// TIA Portal V21 export
// export: Created 2026-11-07T17:04:58.8890969Z, ExportSetting WithDefaults, DisplayName Totally Integrated Automation Portal, DisplayVersion V21, DisplayName STEP 7 Professional, DisplayVersion V21, DisplayName STEP 7 Safety, DisplayVersion V21, DisplayName Tech WebApplication, DisplayVersion V21, DisplayName WinCC Basic/Comfort/Advanced, DisplayVersion V21, DisplayName WinCC Unified, DisplayVersion V21
TextList "TL_Cmd"  ListRange=Decimal
  TextListEntry   EntryType=SingleValue, Text="-"
  TextListEntry   EntryType=SingleValue, From=1, To=1, Text="1 PODIGNI"
  TextListEntry   EntryType=SingleValue, From=2, To=2, Text="2 SPUSTI"
  TextListEntry   EntryType=SingleValue, From=3, To=3, Text="3 POMAKNI"
  TextListEntry   EntryType=SingleValue, From=10, To=10, Text="10 RESET"
